// TIA Portal V21 export
// export: Created 2026-11-10T07:35:02.469601Z, ExportSetting WithDefaults, DisplayName Totally Integrated Automation Portal, DisplayVersion V21 Update 3, DisplayName STEP 7 Professional, DisplayVersion V21 Update 3, DisplayName STEP 7 Safety, DisplayVersion V21, DisplayName Tech WebApplication, DisplayVersion V21, DisplayName WinCC Basic/Comfort/Advanced, DisplayVersion V21 Update 3, DisplayName WinCC Unified, DisplayVersion V21 Update 3
FUNCTION_BLOCK "FB_Lad_ex014"   // FB11, LAD
{ S7_Optimized_Access := 'TRUE' }
VERSION : 0.1
// stored: AutoNumber true, IsIECCheckEnabled false, IsRetainMemResEnabled false, MemoryReserve 100, SetENOAutomatically false, UDAEnableTagReadback false
   VAR_INPUT
      v_nr : RTM;
      v_mode : Byte;
      v_pv : DInt;
      v_ret_val : Int;
   END_VAR
   VAR_OUTPUT
      v_cq : Bool;
      v_cv : DInt;
   END_VAR
BEGIN

REGION Network 1: RTM - Runtime meters
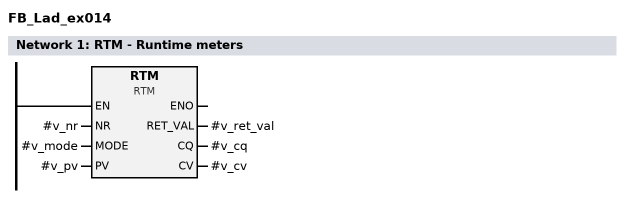
   RUNG wire#powerrail
      { S7_Templates := "nr_type := RTM" } RTM(NR := #v_nr, MODE := #v_mode, PV := #v_pv, RET_VAL => #v_ret_val, CQ => #v_cq, CV => #v_cv)
   END_RUNG
   // the same network as SCL:
   #v_ret_val := RTM(NR := #v_nr, MODE := #v_mode, PV := #v_pv, CQ => #v_cq, CV => #v_cv);
END_REGION
END_FUNCTION_BLOCK
